FUNCTION_BLOCK MOTOR_START_STOP (* Migrated from IEC 61131-3 ST *)
  (* Standard: 61499-2 *)
  (* Version 1.0, 2026-11-06, st2fb *)
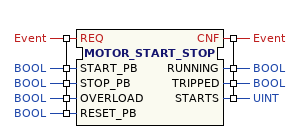
  EVENT_INPUT
    REQ WITH START_PB, STOP_PB, OVERLOAD, RESET_PB;
  END_EVENT
  EVENT_OUTPUT
    CNF WITH RUNNING, TRIPPED, STARTS;
  END_EVENT
  VAR_INPUT
    START_PB : BOOL;
    STOP_PB : BOOL;
    OVERLOAD : BOOL;
    RESET_PB : BOOL;
  END_VAR
  VAR_OUTPUT
    RUNNING : BOOL;
    TRIPPED : BOOL;
    STARTS : UINT;
  END_VAR
  VAR
    PREV_RUNNING : BOOL;
  END_VAR
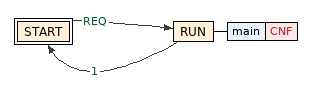
  EC_STATES
    START;
    RUN : main -> CNF;
  END_STATES
  EC_TRANSITIONS
    START TO RUN := REQ;
    RUN TO START := 1;
  END_TRANSITIONS
  ALGORITHM main IN ST:
IF OVERLOAD THEN
  TRIPPED := TRUE;
ELSIF RESET_PB THEN
  TRIPPED := FALSE;
END_IF;
RUNNING := (START_PB OR RUNNING) AND NOT STOP_PB AND NOT TRIPPED;
IF RUNNING AND NOT PREV_RUNNING THEN
  STARTS := STARTS + 1;
END_IF;
PREV_RUNNING := RUNNING;
  END_ALGORITHM
END_FUNCTION_BLOCK
